Fanuc KAREL source: KX00012.KL

PROGRAM KX00012
%NOLOCKGROUP
VAR
  I: INTEGER
  J: INTEGER
  B: BOOLEAN
  F: FILE
  S: STRING[80]
  P: XYZWPR
BEGIN
  UNHOLD
END KX00012
